FUNCTION_BLOCK MOD_Occupation (* Who may command the module. A client first calls the OPC UA method Occupy with a session id it chose; until it calls Release, only commands carrying that session id are accepted. Publishes Occupied (never the id) and tells every block of the module who the owner is. Technical: Module occupation: OPC UA methods Occupy(Session) and Release(Session) answer [Accepted, ErrorID]; publishes Occupied (never the session ID) and shares the owner on a local channel *)
  (* Standard: 61499-2 *)
  (* Version 0.1, 2026-09-28, Project contributors, AAU Smart Production Lab *)
  PACKAGE modlib;
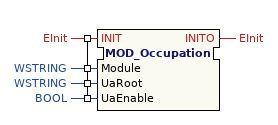
  EVENT_INPUT
    INIT : EInit WITH Module, UaRoot, UaEnable; (* Initialise, once at start-up (the INIT chain); takes the values given with it *)
  END_EVENT
  EVENT_OUTPUT
    INITO : EInit; (* Initialised: the next block of the INIT chain goes on *)
  END_EVENT
  VAR_INPUT
    Module : WSTRING; (* The module's name; its local channels are named after it (loc[<Module>/...]) *)
    UaRoot : WSTRING; (* The module's OPC UA folder, e.g. /Objects/Filling *)
    UaEnable : BOOL; (* Publish on OPC UA *)
  END_VAR
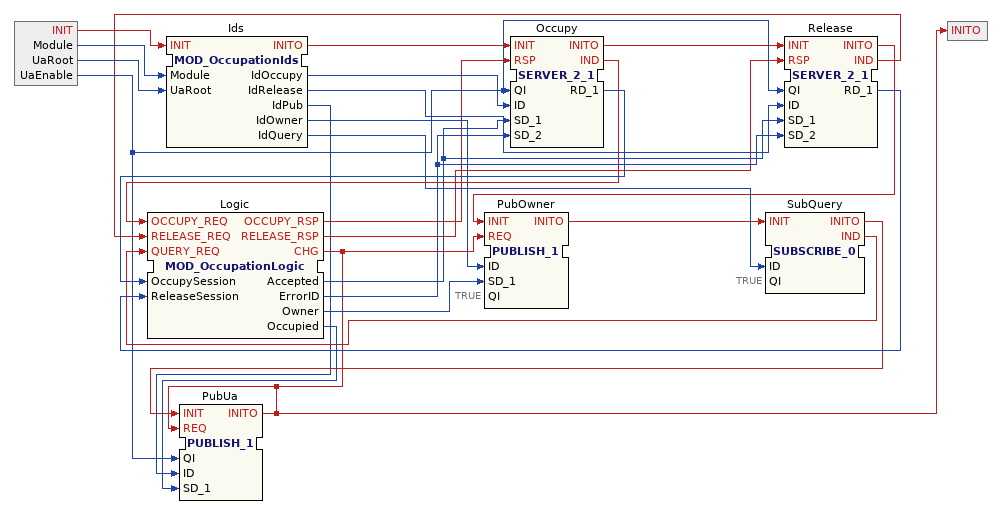
  FBS
    Ids : modlib::MOD_OccupationIds; (* Builds the OPC UA addresses and channel names from the module's name. *)
    Occupy : iec61499::net::SERVER_2_1; (* The OPC UA method Occupation/Occupy(Session). *)
    Release : iec61499::net::SERVER_2_1; (* The OPC UA method Occupation/Release(Session). *)
    Logic : modlib::MOD_OccupationLogic; (* Decides who may occupy and release. *)
    PubOwner : iec61499::net::PUBLISH_1(QI := TRUE); (* Tells every block of the module the owner, on the owner channel. *)
    SubQuery : iec61499::net::SUBSCRIBE_0(QI := TRUE); (* Answers a block that asks who the owner is (at its start). *)
    PubUa : iec61499::net::PUBLISH_1; (* Writes Occupation/Occupied to OPC UA. *)
  END_FBS
  EVENT_CONNECTIONS
    INIT TO Ids.INIT;
    Ids.INITO TO Occupy.INIT;
    Occupy.INITO TO Release.INIT;
    Release.INITO TO PubOwner.INIT;
    PubOwner.INITO TO SubQuery.INIT;
    SubQuery.INITO TO PubUa.INIT;
    PubUa.INITO TO PubUa.REQ;
    PubUa.INITO TO INITO;
    Occupy.IND TO Logic.OCCUPY_REQ;
    Logic.OCCUPY_RSP TO Occupy.RSP;
    Release.IND TO Logic.RELEASE_REQ;
    Logic.RELEASE_RSP TO Release.RSP;
    SubQuery.IND TO Logic.QUERY_REQ;
    Logic.CHG TO PubOwner.REQ;
    Logic.CHG TO PubUa.REQ;
  END_CONNECTIONS
  DATA_CONNECTIONS
    Module TO Ids.Module;
    UaRoot TO Ids.UaRoot;
    UaEnable TO Occupy.QI;
    UaEnable TO Release.QI;
    UaEnable TO PubUa.QI;
    Ids.IdOccupy TO Occupy.ID;
    Ids.IdRelease TO Release.ID;
    Ids.IdPub TO PubUa.ID;
    Ids.IdOwner TO PubOwner.ID;
    Ids.IdQuery TO SubQuery.ID;
    Occupy.RD_1 TO Logic.OccupySession;
    Logic.Accepted TO Occupy.SD_1;
    Logic.ErrorID TO Occupy.SD_2;
    Release.RD_1 TO Logic.ReleaseSession;
    Logic.Accepted TO Release.SD_1;
    Logic.ErrorID TO Release.SD_2;
    Logic.Owner TO PubOwner.SD_1;
    Logic.Occupied TO PubUa.SD_1;
  END_CONNECTIONS
END_FUNCTION_BLOCK
